Staubli VAL3: getMotCount.pgx

public program getMotCount(bool& x_bContain)
  local num l_nI
begin
  x_bContain=false
  for l_nI= 0 to size(nMoveTypeRec)-1
    if nMoveTypeRec[l_nI]!=-1 and nMoveIdRec[l_nI]!=-1
      x_bContain=true
    endIf
  endFor
end
